// TIA Portal V21 export
// export: Created 2026-08-21T20:18:52.4969224Z, ExportSetting None, DisplayName Totally Integrated Automation Portal, DisplayVersion V21, DisplayName STEP 7 Professional, DisplayVersion V21, DisplayName STEP 7 Safety, DisplayVersion V21, DisplayName Tech WebApplication, DisplayVersion V21, DisplayName WinCC Basic/Comfort/Advanced, DisplayVersion V21, DisplayName WinCC Professional, DisplayVersion V21, DisplayName WinCC Unified, DisplayVersion V21
FUNCTION "Service" : Void   // FC11, FBD
TITLE = Service
{ S7_Optimized_Access := 'TRUE' }
AUTHOR : Siemens AG
FAMILY : ServiceControl
VERSION : 1.0
// stored: SetENOAutomatically false
   VAR_TEMP
      ProcedureDone : Bool;
      UnholdingDone : Bool;
      StartingState : Bool;
      CompletingState : Bool;
      PausingState : Bool;
      HoldingState : Bool;
      AbortingState : Bool;
      StoppingState : Bool;
      State : "Service_States";
   END_VAR
   VAR_TEMP   // added for the SCL form of the ladder/FBD networks
      _w1 : Bool;
      _w2 : Bool;
      _w3 : Bool;
      _w4 : Bool;
   END_VAR
BEGIN

REGION Network 1: Parameters and values
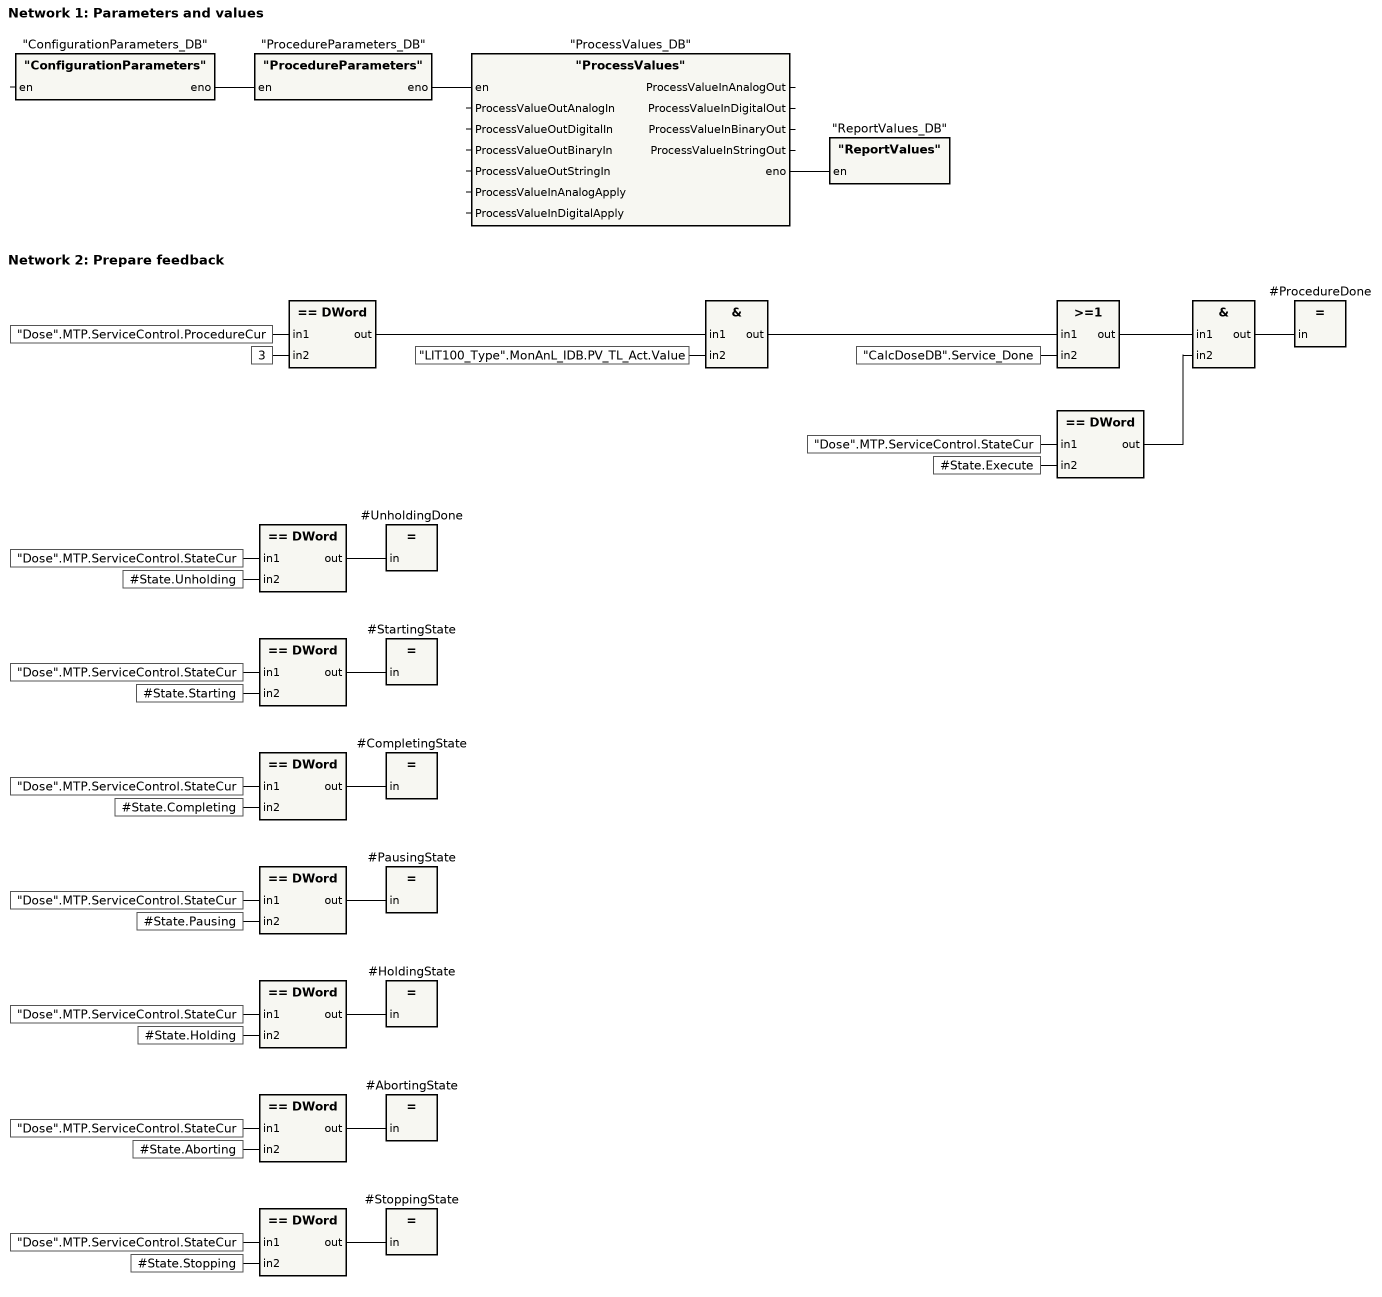
   "ConfigurationParameters_DB"(ENO => #_w1);   // "ConfigurationParameters"
   "ProcedureParameters_DB"(EN := #_w1, ENO => #_w2);   // "ProcedureParameters"
   "ProcessValues_DB"(EN := #_w2, ENO => #_w3);   // "ProcessValues"
   IF #_w3 THEN
       "ReportValues_DB"();   // "ReportValues"
   END_IF;
END_REGION

REGION Network 2: Prepare feedback
   #ProcedureDone := ((("Dose".MTP.ServiceControl.ProcedureCur = 3) AND "LIT100_Type".MonAnL_IDB.PV_TL_Act.Value) OR "CalcDoseDB".Service_Done) AND ("Dose".MTP.ServiceControl.StateCur = #State.Execute);
   #UnholdingDone := "Dose".MTP.ServiceControl.StateCur = #State.Unholding;
   #StartingState := "Dose".MTP.ServiceControl.StateCur = #State.Starting;
   #CompletingState := "Dose".MTP.ServiceControl.StateCur = #State.Completing;
   #PausingState := "Dose".MTP.ServiceControl.StateCur = #State.Pausing;
   #HoldingState := "Dose".MTP.ServiceControl.StateCur = #State.Holding;
   #AbortingState := "Dose".MTP.ServiceControl.StateCur = #State.Aborting;
   #StoppingState := "Dose".MTP.ServiceControl.StateCur = #State.Stopping;
END_REGION

REGION Network 3: Cm P100 feedback
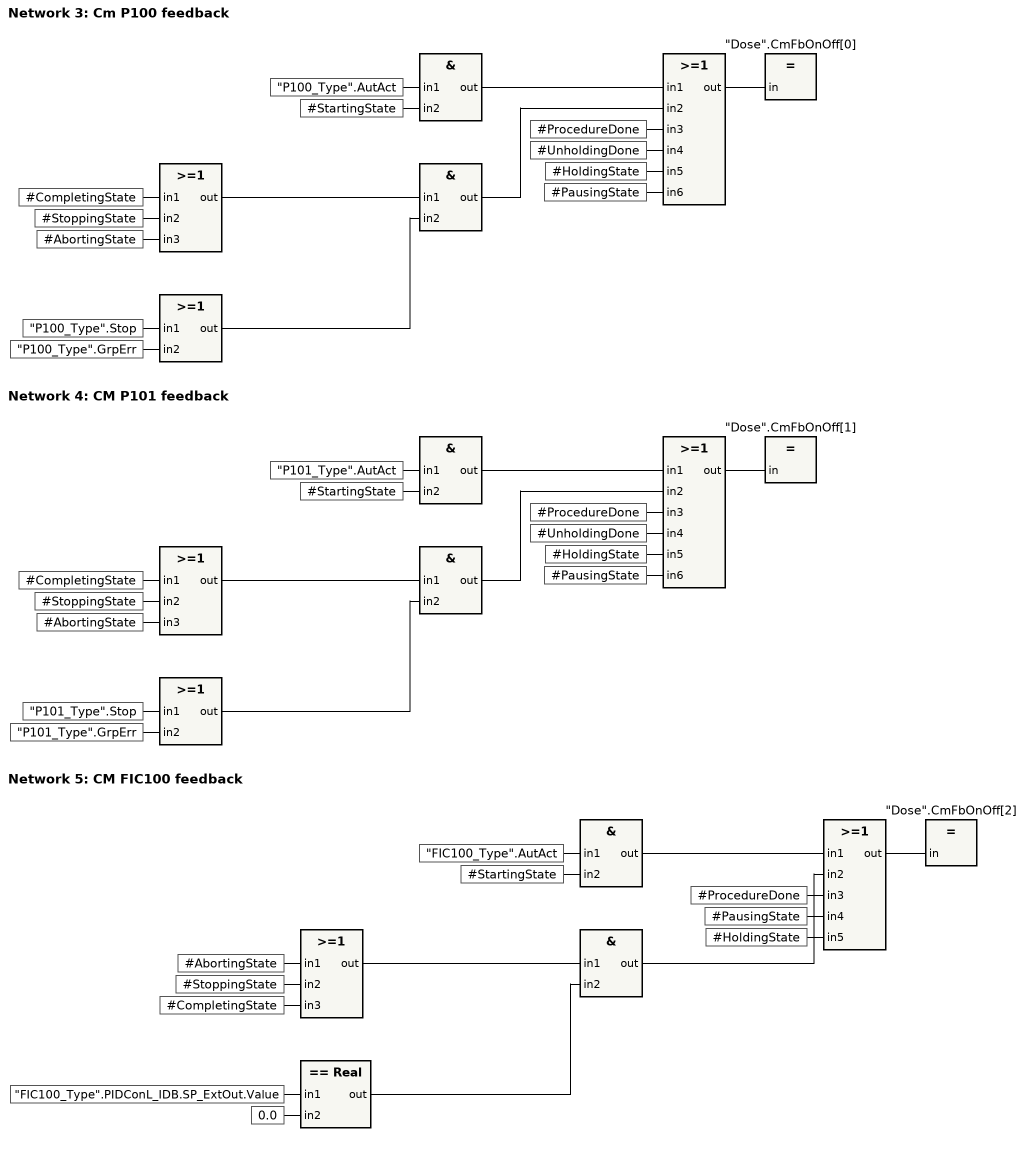
   "Dose".CmFbOnOff[0] := ("P100_Type".AutAct AND #StartingState) OR ((#CompletingState OR #StoppingState OR #AbortingState) AND ("P100_Type".Stop OR "P100_Type".GrpErr)) OR #ProcedureDone OR #UnholdingDone OR #HoldingState OR #PausingState;
END_REGION

REGION Network 4: CM P101 feedback
   "Dose".CmFbOnOff[1] := ("P101_Type".AutAct AND #StartingState) OR ((#CompletingState OR #StoppingState OR #AbortingState) AND ("P101_Type".Stop OR "P101_Type".GrpErr)) OR #ProcedureDone OR #UnholdingDone OR #HoldingState OR #PausingState;
END_REGION

REGION Network 5: CM FIC100 feedback
   "Dose".CmFbOnOff[2] := ("FIC100_Type".AutAct AND #StartingState) OR ((#AbortingState OR #StoppingState OR #CompletingState) AND ("FIC100_Type".PIDConL_IDB.SP_ExtOut.Value = 0.0)) OR #ProcedureDone OR #PausingState OR #HoldingState;
END_REGION

REGION Network 6: CM V100 feedback
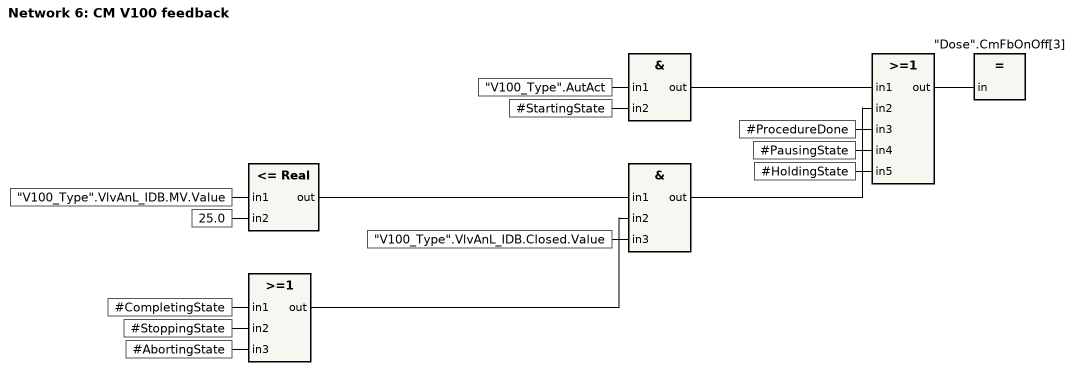
   "Dose".CmFbOnOff[3] := ("V100_Type".AutAct AND #StartingState) OR (("V100_Type".VlvAnL_IDB.MV.Value <= 25.0) AND (#CompletingState OR #StoppingState OR #AbortingState) AND "V100_Type".VlvAnL_IDB.Closed.Value) OR #ProcedureDone OR #PausingState OR #HoldingState;
END_REGION

REGION Network 7: Service
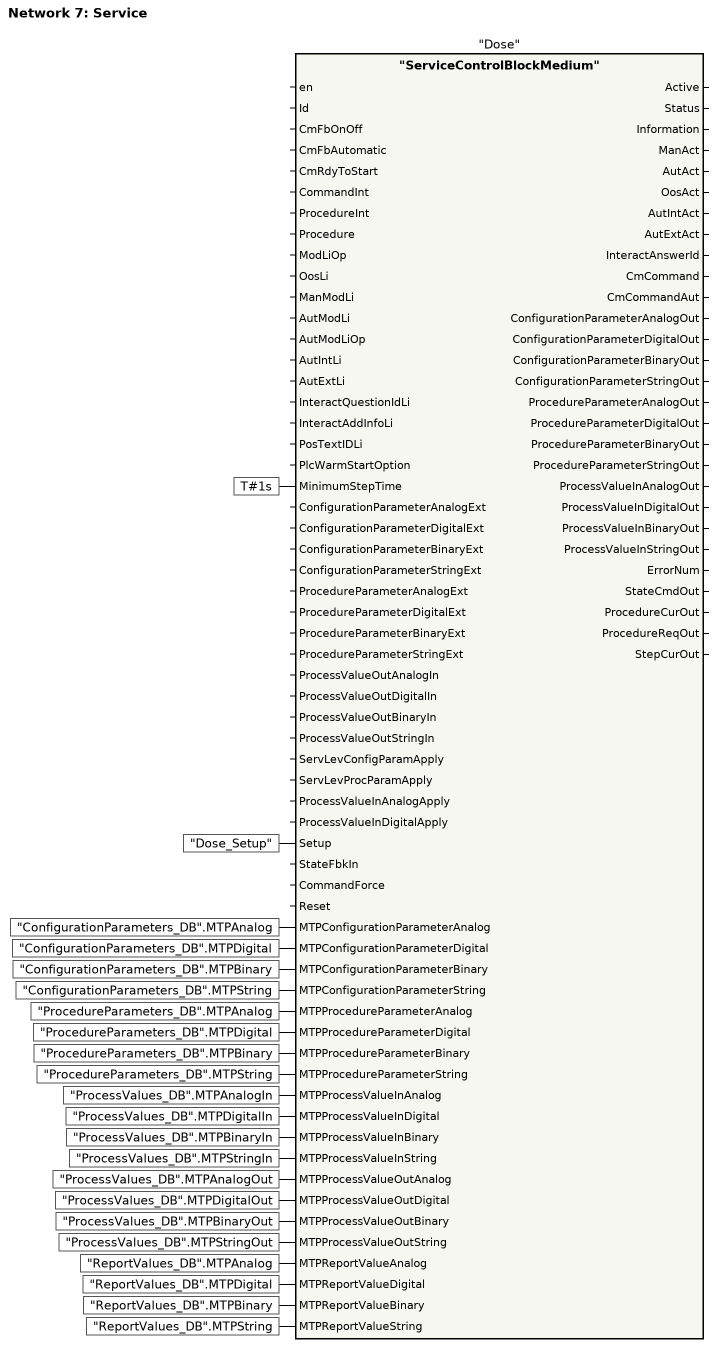
   "Dose"(MinimumStepTime := T#1s,   // "ServiceControlBlockMedium"
          Setup := "Dose_Setup",
          MTPConfigurationParameterAnalog := "ConfigurationParameters_DB".MTPAnalog,
          MTPConfigurationParameterDigital := "ConfigurationParameters_DB".MTPDigital,
          MTPConfigurationParameterBinary := "ConfigurationParameters_DB".MTPBinary,
          MTPConfigurationParameterString := "ConfigurationParameters_DB".MTPString,
          MTPProcedureParameterAnalog := "ProcedureParameters_DB".MTPAnalog,
          MTPProcedureParameterDigital := "ProcedureParameters_DB".MTPDigital,
          MTPProcedureParameterBinary := "ProcedureParameters_DB".MTPBinary,
          MTPProcedureParameterString := "ProcedureParameters_DB".MTPString,
          MTPProcessValueInAnalog := "ProcessValues_DB".MTPAnalogIn,
          MTPProcessValueInDigital := "ProcessValues_DB".MTPDigitalIn,
          MTPProcessValueInBinary := "ProcessValues_DB".MTPBinaryIn,
          MTPProcessValueInString := "ProcessValues_DB".MTPStringIn,
          MTPProcessValueOutAnalog := "ProcessValues_DB".MTPAnalogOut,
          MTPProcessValueOutDigital := "ProcessValues_DB".MTPDigitalOut,
          MTPProcessValueOutBinary := "ProcessValues_DB".MTPBinaryOut,
          MTPProcessValueOutString := "ProcessValues_DB".MTPStringOut,
          MTPReportValueAnalog := "ReportValues_DB".MTPAnalog,
          MTPReportValueDigital := "ReportValues_DB".MTPDigital,
          MTPReportValueBinary := "ReportValues_DB".MTPBinary,
          MTPReportValueString := "ReportValues_DB".MTPString);
END_REGION

REGION Network 8: Service HMI
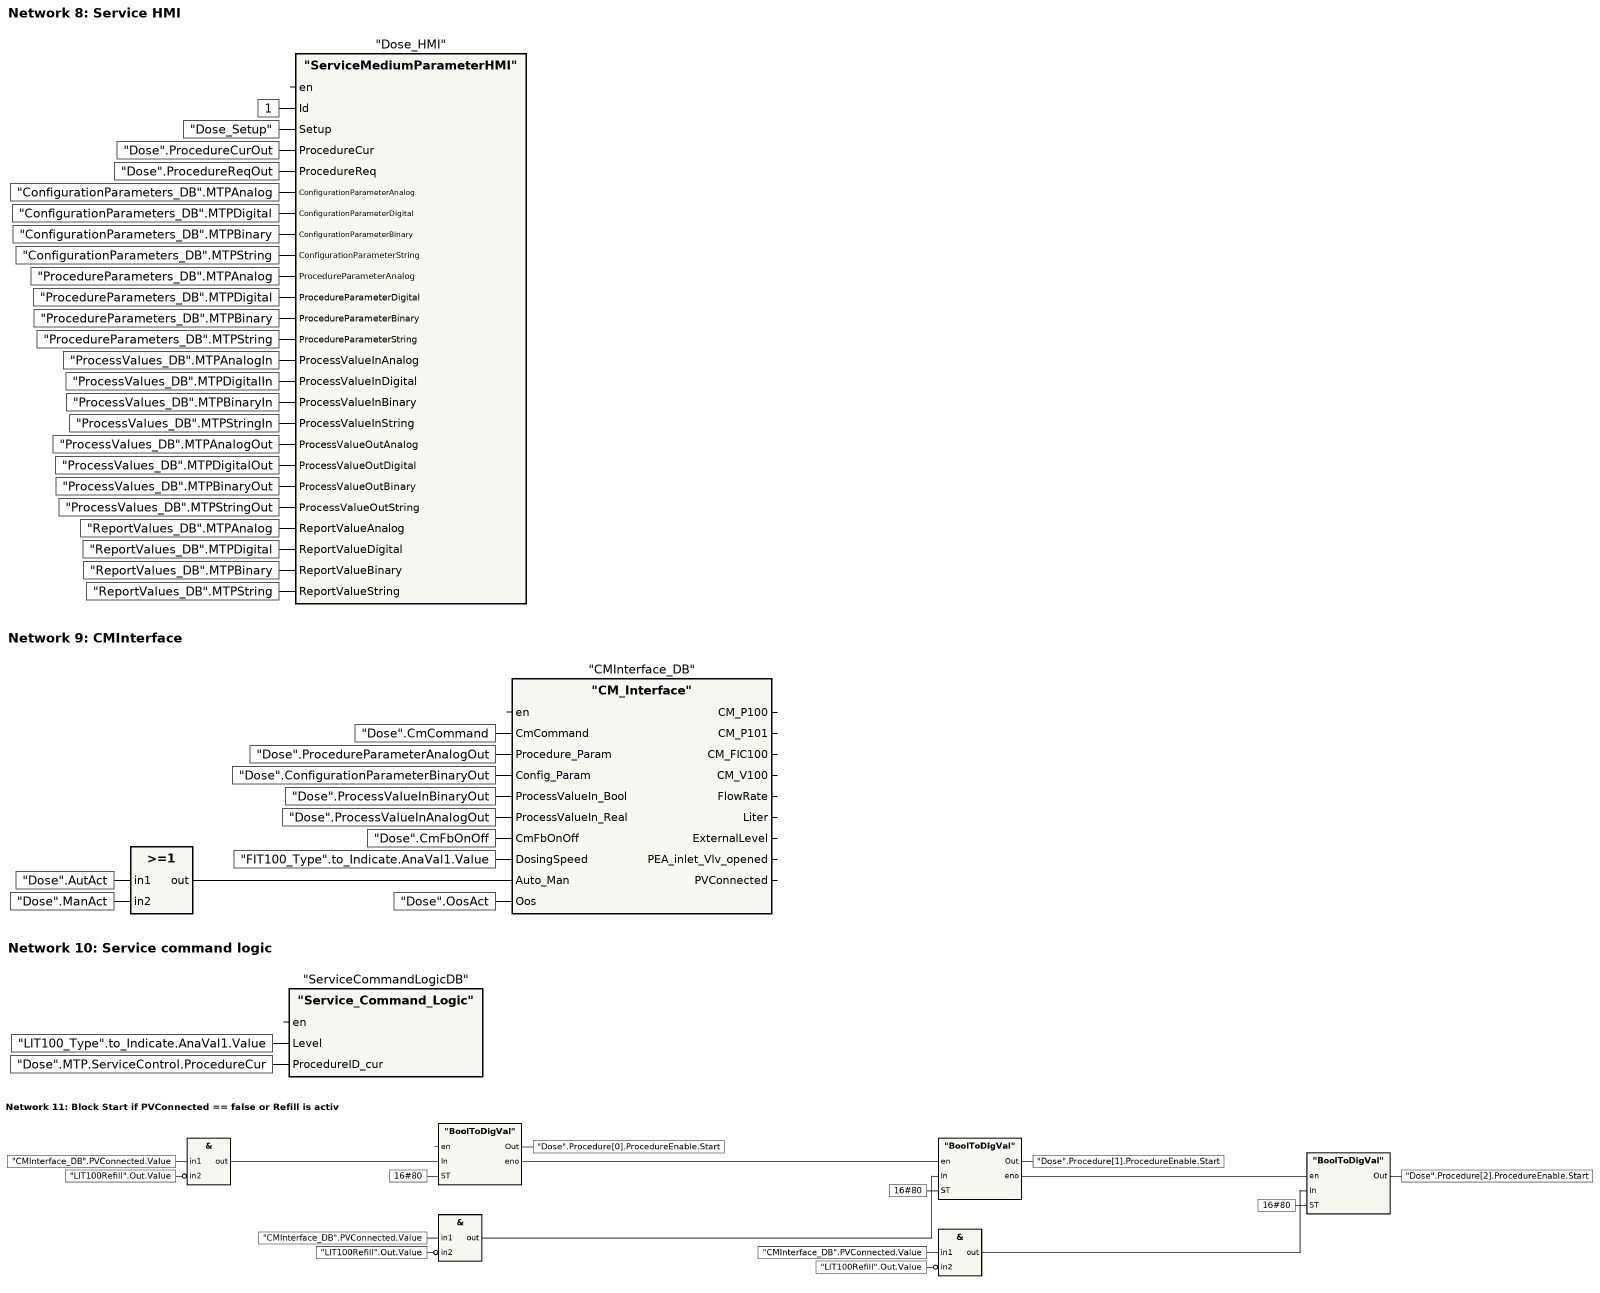
   "Dose_HMI"(Id := 1,   // "ServiceMediumParameterHMI"
              Setup := "Dose_Setup",
              ProcedureCur := "Dose".ProcedureCurOut,
              ProcedureReq := "Dose".ProcedureReqOut,
              ConfigurationParameterAnalog := "ConfigurationParameters_DB".MTPAnalog,
              ConfigurationParameterDigital := "ConfigurationParameters_DB".MTPDigital,
              ConfigurationParameterBinary := "ConfigurationParameters_DB".MTPBinary,
              ConfigurationParameterString := "ConfigurationParameters_DB".MTPString,
              ProcedureParameterAnalog := "ProcedureParameters_DB".MTPAnalog,
              ProcedureParameterDigital := "ProcedureParameters_DB".MTPDigital,
              ProcedureParameterBinary := "ProcedureParameters_DB".MTPBinary,
              ProcedureParameterString := "ProcedureParameters_DB".MTPString,
              ProcessValueInAnalog := "ProcessValues_DB".MTPAnalogIn,
              ProcessValueInDigital := "ProcessValues_DB".MTPDigitalIn,
              ProcessValueInBinary := "ProcessValues_DB".MTPBinaryIn,
              ProcessValueInString := "ProcessValues_DB".MTPStringIn,
              ProcessValueOutAnalog := "ProcessValues_DB".MTPAnalogOut,
              ProcessValueOutDigital := "ProcessValues_DB".MTPDigitalOut,
              ProcessValueOutBinary := "ProcessValues_DB".MTPBinaryOut,
              ProcessValueOutString := "ProcessValues_DB".MTPStringOut,
              ReportValueAnalog := "ReportValues_DB".MTPAnalog,
              ReportValueDigital := "ReportValues_DB".MTPDigital,
              ReportValueBinary := "ReportValues_DB".MTPBinary,
              ReportValueString := "ReportValues_DB".MTPString);
END_REGION

REGION Network 9: CMInterface
   "CMInterface_DB"(CmCommand := "Dose".CmCommand,   // "CM_Interface"
                    Procedure_Param := "Dose".ProcedureParameterAnalogOut,
                    Config_Param := "Dose".ConfigurationParameterBinaryOut,
                    ProcessValueIn_Bool := "Dose".ProcessValueInBinaryOut,
                    ProcessValueIn_Real := "Dose".ProcessValueInAnalogOut,
                    CmFbOnOff := "Dose".CmFbOnOff,
                    DosingSpeed := "FIT100_Type".to_Indicate.AnaVal1.Value,
                    Auto_Man := "Dose".AutAct OR "Dose".ManAct,
                    Oos := "Dose".OosAct);
END_REGION

REGION Network 10: Service command logic
   "ServiceCommandLogicDB"(Level := "LIT100_Type".to_Indicate.AnaVal1.Value,   // "Service_Command_Logic"
                           ProcedureID_cur := "Dose".MTP.ServiceControl.ProcedureCur);
END_REGION

REGION Network 11: Block Start if PVConnected == false or Refill is activ
   "BoolToDigVal"(In := "CMInterface_DB".PVConnected.Value AND NOT "LIT100Refill".Out.Value,
                  ST := 16#80,
                  Out => "Dose".Procedure[0].ProcedureEnable.Start,
                  ENO => #_w1);
   "BoolToDigVal"(EN := #_w1,
                  In := "CMInterface_DB".PVConnected.Value AND NOT "LIT100Refill".Out.Value,
                  ST := 16#80,
                  Out => "Dose".Procedure[1].ProcedureEnable.Start,
                  ENO => #_w2);
   IF #_w2 THEN
       "BoolToDigVal"(In := "CMInterface_DB".PVConnected.Value AND NOT "LIT100Refill".Out.Value,
                      ST := 16#80,
                      Out => "Dose".Procedure[2].ProcedureEnable.Start);
   END_IF;
END_REGION

REGION Network 12: Block Resume and Unholding if refill is activ
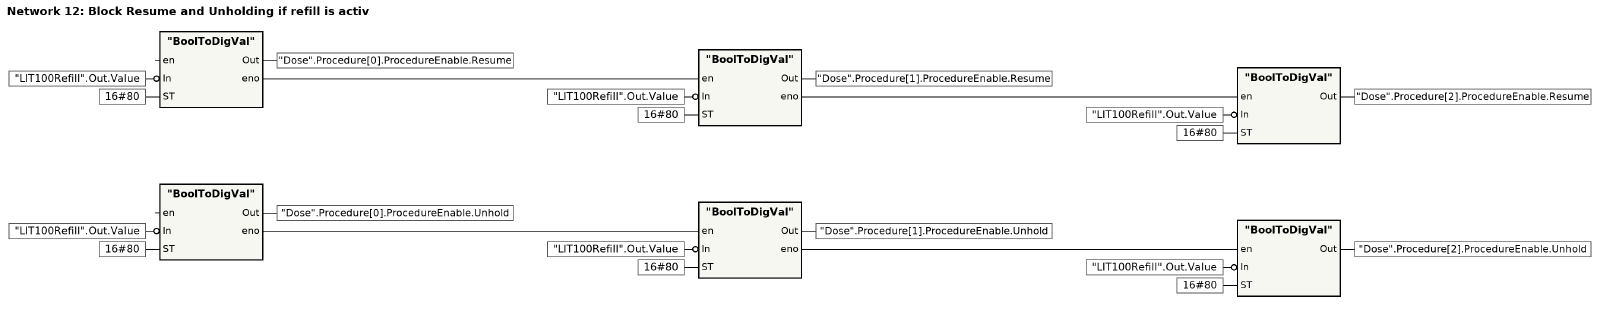
   "BoolToDigVal"(In := NOT "LIT100Refill".Out.Value,
                  ST := 16#80,
                  Out => "Dose".Procedure[0].ProcedureEnable.Resume,
                  ENO => #_w1);
   "BoolToDigVal"(EN := #_w1,
                  In := NOT "LIT100Refill".Out.Value,
                  ST := 16#80,
                  Out => "Dose".Procedure[1].ProcedureEnable.Resume,
                  ENO => #_w2);
   IF #_w2 THEN
       "BoolToDigVal"(In := NOT "LIT100Refill".Out.Value,
                      ST := 16#80,
                      Out => "Dose".Procedure[2].ProcedureEnable.Resume);
   END_IF;
   "BoolToDigVal"(In := NOT "LIT100Refill".Out.Value,
                  ST := 16#80,
                  Out => "Dose".Procedure[0].ProcedureEnable.Unhold,
                  ENO => #_w3);
   "BoolToDigVal"(EN := #_w3,
                  In := NOT "LIT100Refill".Out.Value,
                  ST := 16#80,
                  Out => "Dose".Procedure[1].ProcedureEnable.Unhold,
                  ENO => #_w4);
   IF #_w4 THEN
       "BoolToDigVal"(In := NOT "LIT100Refill".Out.Value,
                      ST := 16#80,
                      Out => "Dose".Procedure[2].ProcedureEnable.Unhold);
   END_IF;
END_REGION

REGION Network 13: Position Text
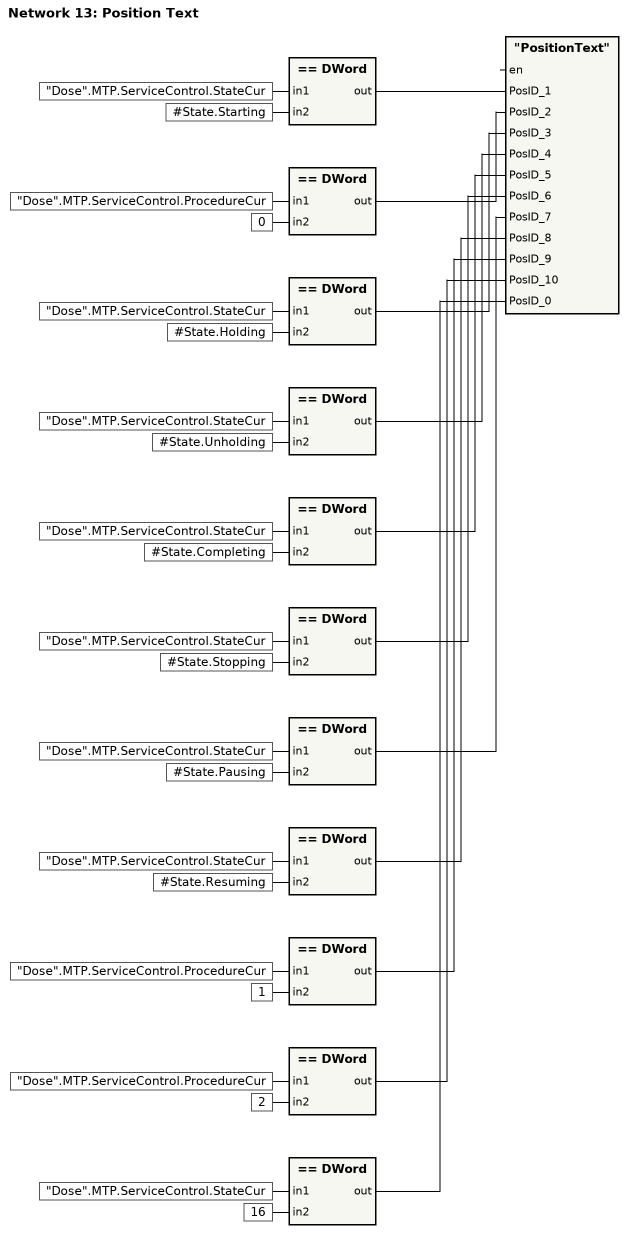
   "PositionText"(PosID_1 := "Dose".MTP.ServiceControl.StateCur = #State.Starting,
                  PosID_2 := "Dose".MTP.ServiceControl.ProcedureCur = 0,
                  PosID_3 := "Dose".MTP.ServiceControl.StateCur = #State.Holding,
                  PosID_4 := "Dose".MTP.ServiceControl.StateCur = #State.Unholding,
                  PosID_5 := "Dose".MTP.ServiceControl.StateCur = #State.Completing,
                  PosID_6 := "Dose".MTP.ServiceControl.StateCur = #State.Stopping,
                  PosID_7 := "Dose".MTP.ServiceControl.StateCur = #State.Pausing,
                  PosID_8 := "Dose".MTP.ServiceControl.StateCur = #State.Resuming,
                  PosID_9 := "Dose".MTP.ServiceControl.ProcedureCur = 1,
                  PosID_10 := "Dose".MTP.ServiceControl.ProcedureCur = 2,
                  PosID_0 := "Dose".MTP.ServiceControl.StateCur = 16);
END_REGION

REGION Network 14: Report values
END_REGION
END_FUNCTION
